// SIMATIC S7-200 project (STEP 7-Micro/WIN), CPU 224 CN REL 02.01

SYMBOL_TABLE USUARIO1
SB_2             I1.2     // Pulsador de paro
SB_1             I1.3     // Pulsador de marcha
QS               I1.4     // Zeta de emergencia
SA               I1.5     // Selector de modo
HL1              Q0.7     // Piloto amarillo
HL2              Q1.0     // Piloto verde
HL3              Q1.1     // Piloto rojo
END_SYMBOL_TABLE

ORGANIZATION_BLOCK PRINCIPAL:OB1
TITLE=COMENTARIOS DEL PROGRAMA
BEGIN
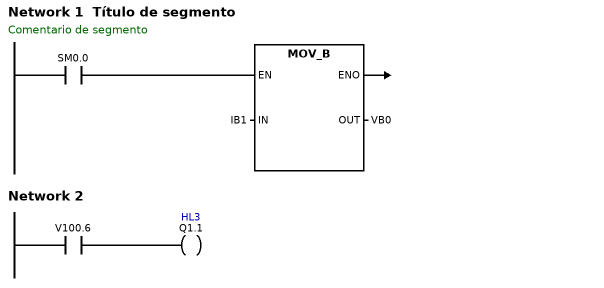
Network 1 // Título de segmento
// Comentario de segmento
LD     SM0.0
MOVB   IB1, VB0
Network 2
LD     V100.6
=      HL3:Q1.1
END_ORGANIZATION_BLOCK
